(* IEC 61131-3 sources: plcassist-cli/packages/volt-lsp-iec/test-corpus/CodesysTestProject/Device/Plc Logic/Application/Library Manager/(unresolved)/systypes interfaces, 1 file *)

(* ---- HANDLECONSTANTS.gvl ---- *)
VAR_GLOBAL
	RTS_INVALID_HANDLE : RTS_IEC_HANDLE := -1;
END_VAR
